(* IEC 61131-3 sources: Repository_IEMA_Test/LMC_PacDrive.device.xml.v3^/Plc Logic.plclogic.xml.v3^/Application.application.xml.v3^/TemplateFullProgrammingFramework/Examples/ExampleDiagSources, 3 files *)

(* ---- FB_ApplicationLoggerDiagSource.fb.st ---- *)
FUNCTION_BLOCK PUBLIC FB_ApplicationLoggerDiagSource
VAR_INPUT
	i_xEnable			: BOOL;
	i_xDiagQuit			: BOOL;
END_VAR

VAR_IN_OUT
	iq_stComStructure	: TPL.ST_DiagnosticsManagerToDiagSource;
END_VAR

VAR_OUTPUT
	q_xActive			: BOOL;
	q_xReady			: BOOL;
	q_etDiag			: GD.ET_Diag := GD.ET_Diag.Ok;
	q_etDiagExt			: ET_DiagExt := ET_DiagExt.Disabled;
	q_sMsg				: STRING[80];
END_VAR

VAR
	xEnableFlag		: BOOL;
	diState			: DINT;

	udiOwnSourceId	: UDINT := 0;

	fbTreeWriter	: TPL.FB_TreeWriter;

	diOldCmd		: DINT := 0;
	diCmdExecState	: DINT := 0;

	etDiagBuffer		: GD.ET_Diag;
	etDiagExtBufferTPL	: TPL.ET_DiagExt;
	etDiagExtBufferAPL	: APL.ET_DiagExt;
	sMsgBuffer			: STRING[80];

	rtrigDiagQuit	: Standard.R_TRIG;

	fbAppLogHandler			: APL.FB_ApplicationLoggerHandler;
	stLogEntry				: APL.ST_LogEntry;
	ifLoggerPoint			: APL.IF_LoggerPoint;
	udiLogEntryCount		: UDINT;
	udiLogEntryCountMax		: UDINT;
	udiLogEntryId			: UDINT;
	udiLoggerPointCount		: UDINT;
	udiLoggerPointCountMax	: UDINT;
END_VAR

VAR CONSTANT
	c_sName			: STRING[TPL.Gc_udiTableWriterMaxNameLength] := 'ApplicationLogger';
	c_sTypeName		: STRING[TPL.Gc_udiTableWriterMaxNameLength] := 'APL_';
END_VAR

IF i_xEnable AND NOT xEnableFlag THEN
	xEnableFlag := TRUE;
	q_xActive := TRUE;
	SetDiagOutputs(	i_etDiag	:= GD.ET_Diag.Ok,
					i_etDiagExt	:= ET_DiagExt.WaitUntilDiagnosticsManagerReady,
					i_sMsg		:= '');
	diState := 10;

ELSIF NOT i_xEnable AND xEnableFlag THEN
	xEnableFlag := FALSE;
	IF udiOwnSourceId <> 0 THEN
		SetDiagOutputs(	i_etDiag	:= GD.ET_Diag.Ok,
						i_etDiagExt	:= ET_DiagExt.WaitUntilDisabled,
						i_sMsg		:= '');
		diState := 100;
	ELSIF udiOwnSourceId = 0 THEN
		SetDiagOutputs(	i_etDiag	:= GD.ET_Diag.Ok,
						i_etDiagExt	:= ET_DiagExt.Disabled,
						i_sMsg		:= '');
	END_IF
END_IF

DiagQuit();

CASE diState OF

	0:	(* Disable & exception state *)
		;

	10:	(* Wait until diagnostics manager ready *)
		IF iq_stComStructure.i_xDiagnosticsManagerReady THEN
			SetDiagOutputs(	i_etDiag	:= GD.ET_Diag.Ok,
							i_etDiagExt	:= ET_DiagExt.WaitUntilDiagSourceRegistered,
							i_sMsg		:= '');
			diState := 20;
		END_IF

	20:	(* Wait until diag source registered *)
		IF NOT iq_stComStructure.i_xDiagnosticsManagerReady THEN
			SetDiagOutputs(	i_etDiag	:= GD.ET_Diag.Ok,
							i_etDiagExt	:= ET_DiagExt.WaitUntilDiagnosticsManagerReady,
							i_sMsg		:= '');
			diState := 10;

		(* only write to register structure if no one else has done it in this cylce *)
		ELSIF (NOT iq_stComStructure.iq_stRegister.xUsed AND iq_stComStructure.iq_stRegister.udiNextId <> 0) THEN
			(* register *)
			iq_stComStructure.iq_stRegister.xUsed := TRUE;
			iq_stComStructure.iq_stRegister.sName		:= c_sName;
			iq_stComStructure.iq_stRegister.sTypeName	:= c_sTypeName;
			udiOwnSourceId := iq_stComStructure.iq_stRegister.udiNextId; (* register with this id; required for the following communication *)

			q_xReady := TRUE;
			SetDiagOutputs(	i_etDiag	:= GD.ET_Diag.Ok,
							i_etDiagExt	:= ET_DiagExt.WaitForCommunication,
							i_sMsg		:= '');
			diState := 30;
		END_IF

	30:	(* Wait for communication *)
		IF NOT iq_stComStructure.i_xDiagnosticsManagerReady THEN

			CancelWriting();

			udiOwnSourceId	:= 0;

			SetDiagOutputs(	i_etDiag	:= GD.ET_Diag.Ok,
							i_etDiagExt	:= ET_DiagExt.WaitUntilDiagnosticsManagerReady,
							i_sMsg		:= '');
			diState := 10;
			RETURN;

		ELSIF (iq_stComStructure.i_udiComWithId = udiOwnSourceId) THEN		(* Am I adressed? *)

			WriteDiagDataControl();

		ELSE
			iq_stComStructure.q_lrProgress := 0.0;

			CancelWriting();

			SetDiagOutputs(	i_etDiag	:= GD.ET_Diag.Ok,
							i_etDiagExt	:= ET_DiagExt.WaitForCommunication,
							i_sMsg		:= '');
		END_IF

	100: (* Wait until disabled *)
		IF NOT iq_stComStructure.i_xDiagnosticsManagerReady THEN

			CancelWriting();

			udiOwnSourceId	:= 0;

			SetDiagOutputs(	i_etDiag	:= GD.ET_Diag.Ok,
							i_etDiagExt	:= ET_DiagExt.Disabled,
							i_sMsg		:= '');

		ELSIF (iq_stComStructure.i_udiComWithId = udiOwnSourceId) THEN		(* Am I adressed? *)

			WriteDiagDataControl();

		(* only write to register structure if no one else has done it in this cylce *)
		ELSIF (NOT iq_stComStructure.iq_stRegister.xUsed AND NOT iq_stComStructure.iq_stRegister.xUnsubscribe) AND
			   NOT iq_stComStructure.i_xDiagnosticsActive THEN

			iq_stComStructure.iq_stRegister.xUsed			:= TRUE;

			iq_stComStructure.iq_stRegister.xUnsubscribe	:= TRUE;
			iq_stComStructure.iq_stRegister.udiSourceId		:= udiOwnSourceId;

			q_xActive := FALSE;

			SetDiagOutputs(	i_etDiag	:= GD.ET_Diag.Ok,
							i_etDiagExt	:= ET_DiagExt.Disabled,
							i_sMsg		:= '');
		END_IF
END_CASE

IF q_xReady THEN
	IF(diCmdExecState <> 0) THEN
		WriteDiagDataToFile();

		IF(iq_stComStructure.iq_diCmd <= 0) THEN
			diOldCmd := iq_stComStructure.iq_diCmd;
		END_IF
	END_IF
END_IF

(* ---- FB_ExampleTableDiagSource.fb.st ---- *)
FUNCTION_BLOCK FB_ExampleTableDiagSource
VAR_INPUT
	i_xEnable			: BOOL;
	i_xDiagQuit			: BOOL;
END_VAR

VAR_IN_OUT
	iq_stComStructure	: TPL.ST_DiagnosticsManagerToDiagSource;
END_VAR

VAR_OUTPUT
	q_xActive			: BOOL;
	q_xReady			: BOOL;
	q_etDiag			: GD.ET_Diag := GD.ET_Diag.Ok;
	q_etDiagExt			: ET_DiagExt := ET_DiagExt.Disabled;
	q_sMsg				: STRING[80];
END_VAR

VAR
	xEnableFlag		: BOOL;
	diState			: DINT;

	udiOwnSourceId : UDINT := 0;

	diOldCmd	: DINT := 0;
	diCmdExecState : DINT := 0;

	fbTableWriter : TPL.FB_TableWriter;

	udiCName : UDINT;
	udiCValue : UDINT;
	udiCC3 : UDINT;

	udiRowCounter : UDINT := 1;

	etDiag			: GD.ET_Diag;
	etDiagExtTPL	: TPL.ET_DiagExt;
	sMsg			: STRING[80];

	rtrigDiagQuit	: Standard.R_TRIG;
END_VAR

VAR CONSTANT
	c_sName : STRING[TPL.Gc_udiTableWriterMaxNameLength] := 'I_am_something';
	c_sTypeName : STRING[TPL.Gc_udiTableWriterMaxNameLength] := 'ExampleTableDiagSource';
	c_udiMaxNumRows : UDINT := 40;
END_VAR

IF i_xEnable AND NOT xEnableFlag THEN
	xEnableFlag := TRUE;

	q_xActive := TRUE;

	SetDiagOutputs(	i_etDiag	:= GD.ET_Diag.Ok,
					i_etDiagExt	:= ET_DiagExt.WaitUntilDiagnosticsManagerReady,
					i_sMsg		:= '');
	diState := 10;

ELSIF NOT i_xEnable AND xEnableFlag THEN
	xEnableFlag := FALSE;

	IF udiOwnSourceId <> 0 THEN
		SetDiagOutputs(	i_etDiag	:= GD.ET_Diag.Ok,
						i_etDiagExt	:= ET_DiagExt.WaitUntilDisabled,
						i_sMsg		:= '');
		diState := 100;

	ELSIF udiOwnSourceId = 0 THEN
		SetDiagOutputs(	i_etDiag	:= GD.ET_Diag.Ok,
						i_etDiagExt	:= ET_DiagExt.Disabled,
						i_sMsg		:= '');
	END_IF
END_IF

DiagQuit();

CASE diState OF

	0:	(* Disable & exception state *)

	10:	(* Wait until diagnostics manager ready *)
		IF iq_stComStructure.i_xDiagnosticsManagerReady THEN

			SetDiagOutputs(	i_etDiag	:= GD.ET_Diag.Ok,
							i_etDiagExt	:= ET_DiagExt.WaitUntilDiagSourceRegistered,
							i_sMsg		:= '');
			diState := 20;
		END_IF

	20:	(* Wait until diag source registered *)
		IF NOT iq_stComStructure.i_xDiagnosticsManagerReady THEN

			SetDiagOutputs(	i_etDiag	:= GD.ET_Diag.Ok,
							i_etDiagExt	:= ET_DiagExt.WaitUntilDiagnosticsManagerReady,
							i_sMsg		:= '');
			diState := 10;
			RETURN;

		(* only write to register structure if no one else has done it in this cylce *)
		ELSIF (NOT iq_stComStructure.iq_stRegister.xUsed AND iq_stComStructure.iq_stRegister.udiNextId <> 0) THEN
			(* register *)
			iq_stComStructure.iq_stRegister.xUsed := TRUE;

			iq_stComStructure.iq_stRegister.sName		:= c_sName;
			iq_stComStructure.iq_stRegister.sTypeName	:= c_sTypeName;

			udiOwnSourceId := iq_stComStructure.iq_stRegister.udiNextId; (* register with this id; required for the following communication *)
		ELSE
			RETURN;
		END_IF

		q_xReady := TRUE;

		SetDiagOutputs(	i_etDiag	:= GD.ET_Diag.Ok,
						i_etDiagExt	:= ET_DiagExt.WaitForCommunication,
						i_sMsg		:= '');
		diState := 30;

	30:	(* Wait for communication *)
		IF NOT iq_stComStructure.i_xDiagnosticsManagerReady THEN

			CancelWriting();

			udiOwnSourceId	:= 0;

			SetDiagOutputs(	i_etDiag	:= GD.ET_Diag.Ok,
							i_etDiagExt	:= ET_DiagExt.WaitUntilDiagnosticsManagerReady,
							i_sMsg		:= '');
			diState := 10;
			RETURN;

		ELSIF (iq_stComStructure.i_udiComWithId = udiOwnSourceId) THEN		(* Am I adressed? *)

			WriteDiagDataControl();

		ELSE
			iq_stComStructure.q_lrProgress := 0.0;

			CancelWriting();

			SetDiagOutputs(	i_etDiag	:= GD.ET_Diag.Ok,
							i_etDiagExt	:= ET_DiagExt.WaitForCommunication,
							i_sMsg		:= '');
		END_IF

	100: (* Wait until disabled *)
		IF NOT iq_stComStructure.i_xDiagnosticsManagerReady THEN

			CancelWriting();

			udiOwnSourceId	:= 0;

			SetDiagOutputs(	i_etDiag	:= GD.ET_Diag.Ok,
							i_etDiagExt	:= ET_DiagExt.Disabled,
							i_sMsg		:= '');

		ELSIF (iq_stComStructure.i_udiComWithId = udiOwnSourceId) THEN		(* Am I adressed? *)

			WriteDiagDataControl();

		(* only write to register structure if no one else has done it in this cylce *)
		ELSIF (NOT iq_stComStructure.iq_stRegister.xUsed AND NOT iq_stComStructure.iq_stRegister.xUnsubscribe) AND
			   NOT iq_stComStructure.i_xDiagnosticsActive THEN

			iq_stComStructure.iq_stRegister.xUsed			:= TRUE;

			iq_stComStructure.iq_stRegister.xUnsubscribe	:= TRUE;
			iq_stComStructure.iq_stRegister.udiSourceId		:= udiOwnSourceId;

			q_xActive := FALSE;

			SetDiagOutputs(	i_etDiag	:= GD.ET_Diag.Ok,
							i_etDiagExt	:= ET_DiagExt.Disabled,
							i_sMsg		:= '');
		END_IF
END_CASE

IF q_xActive THEN
	IF(diCmdExecState <> 0) THEN
		WriteDiagDataToFile();

		IF(iq_stComStructure.iq_diCmd <= 0) THEN
			diOldCmd := iq_stComStructure.iq_diCmd;
		END_IF
	END_IF
END_IF

(* ---- FB_ExampleTreeDiagSource.fb.st ---- *)
FUNCTION_BLOCK FB_ExampleTreeDiagSource
VAR_INPUT
	i_xEnable			: BOOL;
	i_xDiagQuit			: BOOL;
END_VAR

VAR_IN_OUT
	iq_stComStructure	: TPL.ST_DiagnosticsManagerToDiagSource;
END_VAR

VAR_OUTPUT
	q_xActive			: BOOL;
	q_xReady			: BOOL;
	q_etDiag			: GD.ET_Diag := GD.ET_Diag.Ok;
	q_etDiagExt			: ET_DiagExt := ET_DiagExt.Disabled;
	q_sMsg				: STRING[80];
END_VAR

VAR
	xEnableFlag		: BOOL;
	diState			: DINT;

	udiOwnSourceId : UDINT := 0;

	fbTreeWriter	: TPL.FB_TreeWriter;

	diOldCmd	: DINT := 0;
	diCmdExecState : DINT := 0;

	uiMaxNodePerLevel : UINT := 7;

	uiLevelCounter : UINT := 1;
	auiNodeCounter : ARRAY[1..c_uiMaxLevel] OF UINT;
	uiNodeId : UINT := 1;
	lrSumNodes : LREAL := 1;

	uiTmp : UINT := 0;

	etDiag			: GD.ET_Diag;
	etDiagExtTPL	: TPL.ET_DiagExt;
	sMsg			: STRING[80];

	rtrigDiagQuit	: Standard.R_TRIG;
END_VAR

VAR CONSTANT
	c_sName : STRING[TPL.Gc_udiTableWriterMaxNameLength] := 'I_am_a_Tree';
	c_sTypeName : STRING[TPL.Gc_udiTableWriterMaxNameLength] := 'ExampleTreeDiagSource';
	c_uiMaxLevel : UINT := 5;
END_VAR

IF i_xEnable AND NOT xEnableFlag THEN
	xEnableFlag := TRUE;

	q_xActive := TRUE;

	SetDiagOutputs(	i_etDiag	:= GD.ET_Diag.Ok,
					i_etDiagExt	:= ET_DiagExt.WaitUntilDiagnosticsManagerReady,
					i_sMsg		:= '');
	diState := 10;

ELSIF NOT i_xEnable AND xEnableFlag THEN
	xEnableFlag := FALSE;

	IF udiOwnSourceId <> 0 THEN
		SetDiagOutputs(	i_etDiag	:= GD.ET_Diag.Ok,
						i_etDiagExt	:= ET_DiagExt.WaitUntilDisabled,
						i_sMsg		:= '');
		diState := 100;

	ELSIF udiOwnSourceId = 0 THEN
		SetDiagOutputs(	i_etDiag	:= GD.ET_Diag.Ok,
						i_etDiagExt	:= ET_DiagExt.Disabled,
						i_sMsg		:= '');
	END_IF
END_IF

DiagQuit();

CASE diState OF

	0:	(* Disable & exception state *)

	10:	(* Wait until diagnostics manager ready *)
		IF iq_stComStructure.i_xDiagnosticsManagerReady THEN

			SetDiagOutputs(	i_etDiag	:= GD.ET_Diag.Ok,
							i_etDiagExt	:= ET_DiagExt.WaitUntilDiagSourceRegistered,
							i_sMsg		:= '');
			diState := 20;
		END_IF

	20:	(* Wait until diag source registered *)
		IF NOT iq_stComStructure.i_xDiagnosticsManagerReady THEN

			SetDiagOutputs(	i_etDiag	:= GD.ET_Diag.Ok,
							i_etDiagExt	:= ET_DiagExt.WaitUntilDiagnosticsManagerReady,
							i_sMsg		:= '');
			diState := 10;
			RETURN;

		(* only write to register structure if no one else has done it in this cylce *)
		ELSIF (NOT iq_stComStructure.iq_stRegister.xUsed AND iq_stComStructure.iq_stRegister.udiNextId <> 0) THEN
			(* register *)
			iq_stComStructure.iq_stRegister.xUsed := TRUE;

			iq_stComStructure.iq_stRegister.sName		:= c_sName;
			iq_stComStructure.iq_stRegister.sTypeName	:= c_sTypeName;

			udiOwnSourceId := iq_stComStructure.iq_stRegister.udiNextId; (* register with this id; required for the following communication *)
		ELSE
			RETURN;
		END_IF

		q_xReady := TRUE;

		SetDiagOutputs(	i_etDiag	:= GD.ET_Diag.Ok,
						i_etDiagExt	:= ET_DiagExt.WaitForCommunication,
						i_sMsg		:= '');
		diState := 30;

	30:	(* Wait for communication *)
		IF NOT iq_stComStructure.i_xDiagnosticsManagerReady THEN

			CancelWriting();

			udiOwnSourceId	:= 0;

			SetDiagOutputs(	i_etDiag	:= GD.ET_Diag.Ok,
							i_etDiagExt	:= ET_DiagExt.WaitUntilDiagnosticsManagerReady,
							i_sMsg		:= '');
			diState := 10;
			RETURN;

		ELSIF (iq_stComStructure.i_udiComWithId = udiOwnSourceId) THEN		(* Am I adressed? *)

			WriteDiagDataControl();

		ELSE
			iq_stComStructure.q_lrProgress := 0.0;

			CancelWriting();

			SetDiagOutputs(	i_etDiag	:= GD.ET_Diag.Ok,
							i_etDiagExt	:= ET_DiagExt.WaitForCommunication,
							i_sMsg		:= '');
		END_IF

	100: (* Wait until disabled *)
		IF NOT iq_stComStructure.i_xDiagnosticsManagerReady THEN

			CancelWriting();

			udiOwnSourceId	:= 0;

			SetDiagOutputs(	i_etDiag	:= GD.ET_Diag.Ok,
							i_etDiagExt	:= ET_DiagExt.Disabled,
							i_sMsg		:= '');

		ELSIF (iq_stComStructure.i_udiComWithId = udiOwnSourceId) THEN		(* Am I adressed? *)

			WriteDiagDataControl();

		(* only write to register structure if no one else has done it in this cylce *)
		ELSIF (NOT iq_stComStructure.iq_stRegister.xUsed AND NOT iq_stComStructure.iq_stRegister.xUnsubscribe) AND
			   NOT iq_stComStructure.i_xDiagnosticsActive THEN

			iq_stComStructure.iq_stRegister.xUsed			:= TRUE;

			iq_stComStructure.iq_stRegister.xUnsubscribe	:= TRUE;
			iq_stComStructure.iq_stRegister.udiSourceId		:= udiOwnSourceId;

			q_xActive := FALSE;

			SetDiagOutputs(	i_etDiag	:= GD.ET_Diag.Ok,
							i_etDiagExt	:= ET_DiagExt.Disabled,
							i_sMsg		:= '');
		END_IF
END_CASE

IF q_xActive THEN
	IF(diCmdExecState <> 0) THEN
		WriteDiagDataToFile();

		IF(iq_stComStructure.iq_diCmd <= 0) THEN
			diOldCmd := iq_stComStructure.iq_diCmd;
		END_IF
	END_IF
END_IF
